Universal Robots URScript: T004_mistralai_Mistral-Large-3-675B-Instruct-2512-NVFP4_edit_perf_rep1.urscript

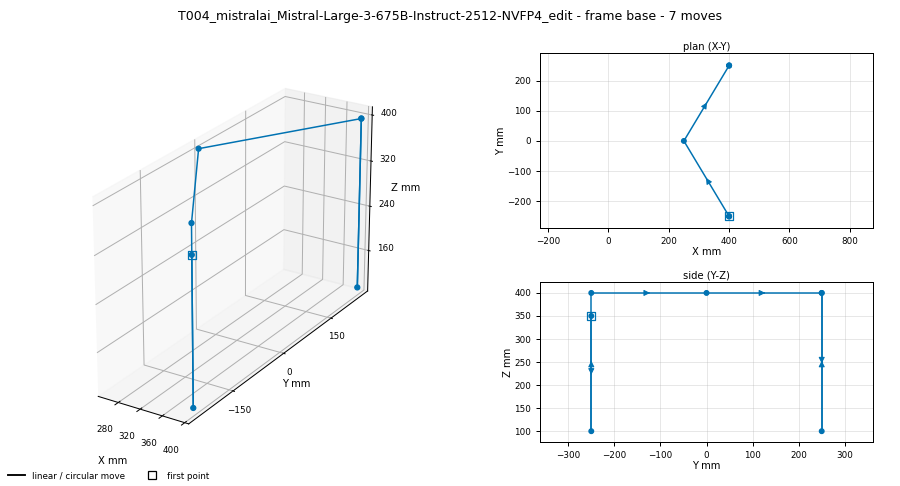
[picture p0: tool path of T004_mistralai_Mistral-Large-3-675B-Instruct-2512-NVFP4_edit_perf_rep1.urscript in frame base, 7 of 9 moves have a stored position in this frame; points joined in program order, loops and branches not executed]
# Task: T004 — Optimized Multi-waypoint SSM pick-place with obstacle avoidance
# Operating mode: collaborative | Max TCP speed: 0.250 m/s
# Robot: ur5e | Payload: 1.5 kg

def task_T004():
  # [0] Verify E-Stop clear
  if (get_digital_in(0) == True):
    popup("E-Stop active — aborting program.", error=True)
    halt
  end

  # [1] Home position - increased acceleration
  movej([0.0000, -1.5708, 1.5708, -1.5708, -1.5708, 0.0000], a=2.0000, v=1.0000)

  # [2] WP1 — Above pick station - increased speed and acceleration
  movel(p[0.400000, -0.250000, 0.350000, 0.0000, 3.1416, 0.0000], a=1.2000, v=0.2500, r=0.0150)

  # [3] WP2 — Descend to pick - optimized acceleration
  movel(p[0.400000, -0.250000, 0.100000, 0.0000, 3.1416, 0.0000], a=0.8000, v=0.1500)

  # [4] Gripper CLOSE
  set_digital_out(0, True)

  # [5] Grip settle - reduced time
  sleep(0.1000)

  # [6] WP3 — Lift above pick - increased speed and acceleration
  movel(p[0.400000, -0.250000, 0.400000, 0.0000, 3.1416, 0.0000], a=1.2000, v=0.2500, r=0.0200)

  # [7] WP4 — Obstacle avoidance waypoint - increased speed and acceleration
  movel(p[0.250000, 0.000000, 0.400000, 0.0000, 3.1416, 0.0000], a=1.2000, v=0.2500, r=0.0300)

  # [8] WP5 — Above place station - increased speed and acceleration
  movel(p[0.400000, 0.250000, 0.400000, 0.0000, 3.1416, 0.0000], a=1.2000, v=0.2500, r=0.0200)

  # [9] WP6 — Descend to place - optimized acceleration
  movel(p[0.400000, 0.250000, 0.100000, 0.0000, 3.1416, 0.0000], a=0.8000, v=0.1500)

  # [10] Gripper OPEN
  set_digital_out(0, False)

  # [11] Release settle - reduced time
  sleep(0.1000)

  # [12] WP7 — Retract above place - increased speed and acceleration
  movel(p[0.400000, 0.250000, 0.400000, 0.0000, 3.1416, 0.0000], a=1.2000, v=0.2500, r=0.0100)

  # [13] Return to home - increased speed and acceleration
  movej([0.0000, -1.5708, 1.5708, -1.5708, -1.5708, 0.0000], a=2.0000, v=1.0000)

end

# Entry point
task_T004()
